SUBAPPLICATION AX_SUBSCRIBE_BG3_WEB_Option_OPC (* OPC-UA Remote-Subscribe + VT-Hintergrundfarbe auf SoftKey UND AuxFunction2 + lokaler Web-Republish - Option-Lib-Variante von AX_SUBSCRIBE_BG3_WEB_OPC: AX_SUBSCRIBE_1, STATUS_WEB_PUBLISH UND GreenWhiteBackground3_AX (hat seit dem QI/QO-Rollout echtes QI/QO) werden vom Option::AOption-Socket initialisiert und gated - Subscribe/Publish sequenziell, GreenWhiteBackground3_AX parallel dazu (E_REND_2_INITO wartet auf beide Zweige, sonst verliert der erste Remote-Wert das Rennen gegen die eigene Q_BackgroundColour-Initialisierung). AOption_OUT reicht die Aktivierung an eine nachgeschaltete Gruppe weiter (Daisy-Chain). *)
  (* Standard: 61499-2; Description: Copyright (c) 2026 Büngener Schuder GmbH This program and the accompanying materials are made available under the terms of the Eclipse Public License 2.0 which is available at https://www.eclipse.org/legal/epl-2.0/ SPDX-License-Identifier: EPL-2.0 *)
  (* Version 1.2, 2026-10-30, Franz Höpfinger, Büngener Schuder GmbH, Remote-Clients mit Remote_Init_Retry: Kette (und Option-INIT_CNF) wartet nicht mehr auf die Gegenstation, nach INITO- neuer Versuch nach 2 s (forte #1092, sonst 60 s pro fehlendem Node und danach tot). *)
  (* Version 1.1, 2026-10-15, Franz Höpfinger, Büngener Schuder GmbH, GreenWhiteBackground3_AX jetzt mitgegated (hat seit QI/QO-Rollout echtes QI/QO, v1.0-Annahme war veraltet) - behebt 'Softkey da, aber Hintergrund reagiert nicht'. E_REND_2_INITO ergaenzt: GreenWhiteBackground3_AX.INIT parallel statt sequenziell nach STATUS_WEB_PUBLISH, sonst verliert der erste eintreffende Remote-Wert das Rennen gegen die eigene Q_BackgroundColour-Init (behebt Folgeregression 'Umschaltung passt, Farbe nicht'). *)
  (* Version 1.0, 2026-10-13, Franz Höpfinger, Büngener Schuder GmbH, initial implementation - Option-Lib-Variante von AX_SUBSCRIBE_BG3_WEB_OPC, nur fuer Softkey_Aux_IXA_TO_Remote_WRITE_BG_Option_OPC gebaut (Status-Haelfte). Bewusst NICHT alle Bausteine gegated - nur die mit echtem QI (AX_SUBSCRIBE_1, STATUS_WEB_PUBLISH), GreenWhiteBackground3_AX bleibt wie im Original unangetastet. *)
  PACKAGE MyLib::sys;
  IMPORT isobus::UT::Q::const::IDs::ID_NULL;
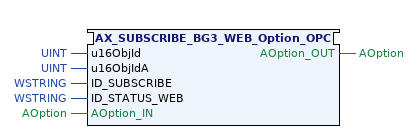
  VAR_INPUT
    u16ObjId : UINT := ID_NULL; (* Object ID SoftKey/Hintergrund (VT) *)
    u16ObjIdA : UINT := ID_NULL; (* Object ID AuxFunction2/Hintergrund (VT) *)
    ID_SUBSCRIBE : WSTRING; (* Remote-Subscribe-Adresse (Status/Farbe, ACTION=SUBSCRIBE) *)
    ID_STATUS_WEB : WSTRING; (* Lokale Publish-Adresse (auf diesem Modul) fuer den vom Zielmodul zurueckgemeldeten Zustand - damit ein Web-Client (z.B. vt-ui-mirror) dieselbe Hintergrundfarbe wie das echte VT zeigen kann *)
  END_VAR
  SOCKETS
    AOption_IN : Option::AOption; (* Treibt INIT/QI von AX_SUBSCRIBE_1/STATUS_WEB_PUBLISH - typischerweise von Softkey_Aux_IXA_TO_Remote_WRITE_Option.AOption_OUT (derselbe Options-Kanal, sequenziell nach der Kommando-Seite) *)
  END_SOCKETS
  PLUGS
    AOption_OUT : Option::AOption; (* Reicht die Aktivierung an eine nachgeschaltete Gruppe weiter (Daisy-Chain) - unbenutzt lassen, wenn nichts weiter folgt *)
  END_PLUGS
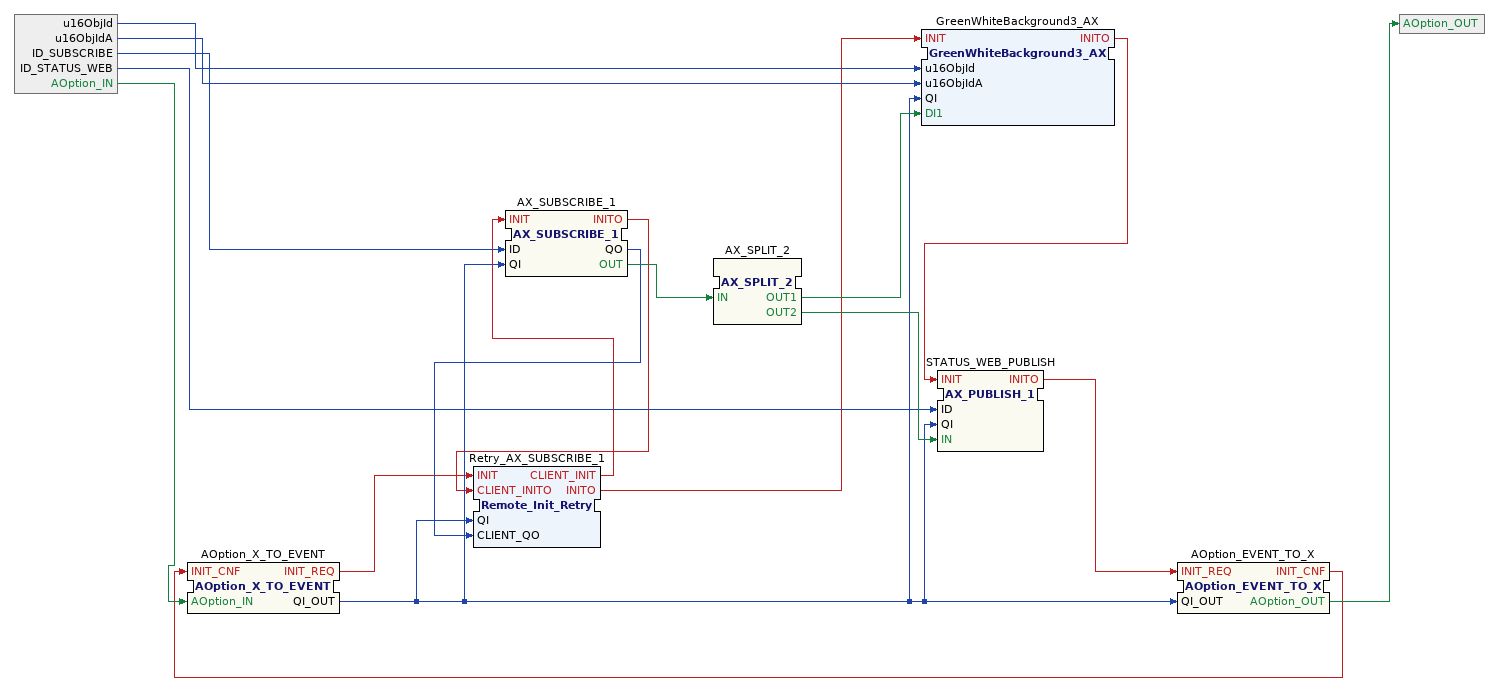
  FBS
    AX_SUBSCRIBE_1 : adapter::net::AX_SUBSCRIBE_1;
    AX_SPLIT_2 : adapter::events::unidirectional::AX_SPLIT_2;
    STATUS_WEB_PUBLISH : adapter::net::AX_PUBLISH_1;
    AOption_X_TO_EVENT : Option::conversion::AOption_X_TO_EVENT;
    AOption_EVENT_TO_X : Option::conversion::AOption_EVENT_TO_X;
  END_FBS
  SUBAPPS
    GreenWhiteBackground3_AX : MyLib::sys::GreenWhiteBackground3_AX;
    Retry_AX_SUBSCRIBE_1 : MyLib::sys::Remote_Init_Retry;
  END_SUBAPPS
  EVENT_CONNECTIONS
    AOption_X_TO_EVENT.INIT_REQ TO Retry_AX_SUBSCRIBE_1.INIT;
    Retry_AX_SUBSCRIBE_1.CLIENT_INIT TO AX_SUBSCRIBE_1.INIT;
    AX_SUBSCRIBE_1.INITO TO Retry_AX_SUBSCRIBE_1.CLIENT_INITO;
    Retry_AX_SUBSCRIBE_1.INITO TO GreenWhiteBackground3_AX.INIT;
    GreenWhiteBackground3_AX.INITO TO STATUS_WEB_PUBLISH.INIT;
    STATUS_WEB_PUBLISH.INITO TO AOption_EVENT_TO_X.INIT_REQ;
    AOption_EVENT_TO_X.INIT_CNF TO AOption_X_TO_EVENT.INIT_CNF;
  END_CONNECTIONS
  DATA_CONNECTIONS
    AOption_X_TO_EVENT.QI_OUT TO Retry_AX_SUBSCRIBE_1.QI;
    AX_SUBSCRIBE_1.QO TO Retry_AX_SUBSCRIBE_1.CLIENT_QO;
    u16ObjId TO GreenWhiteBackground3_AX.u16ObjId;
    u16ObjIdA TO GreenWhiteBackground3_AX.u16ObjIdA;
    ID_SUBSCRIBE TO AX_SUBSCRIBE_1.ID;
    ID_STATUS_WEB TO STATUS_WEB_PUBLISH.ID;
    AOption_X_TO_EVENT.QI_OUT TO AX_SUBSCRIBE_1.QI;
    AOption_X_TO_EVENT.QI_OUT TO STATUS_WEB_PUBLISH.QI;
    AOption_X_TO_EVENT.QI_OUT TO GreenWhiteBackground3_AX.QI;
    AOption_X_TO_EVENT.QI_OUT TO AOption_EVENT_TO_X.QI_OUT;
  END_CONNECTIONS
  ADAPTER_CONNECTIONS
    AX_SUBSCRIBE_1.OUT TO AX_SPLIT_2.IN;
    AX_SPLIT_2.OUT1 TO GreenWhiteBackground3_AX.DI1;
    AX_SPLIT_2.OUT2 TO STATUS_WEB_PUBLISH.IN;
    AOption_IN TO AOption_X_TO_EVENT.AOption_IN;
    AOption_EVENT_TO_X.AOption_OUT TO AOption_OUT;
  END_CONNECTIONS
END_SUBAPPLICATION
